Staubli VAL3: teachPoint1.pgx

public program teachPoint1(string x_sKey, num x_nIndex, num x_nPointIndex)
  local num l_nFrameIndex
  local num l_nToolIndex
  local frame l_fFrame
  local tool l_tTool
  local bool l_bResult
  local pointRx l_pPoint
begin
  link(l_tTool,flange)
  link(l_fFrame,world)
  //  l_bResult=userPageConfirm("是否记录当前点位："+toString("",x_nIndex))
  //  if l_bResult
  l_nFrameIndex=trajTemp:tTrajItem[x_sKey].nFrameIndex
  l_nToolIndex=trajTemp:tTrajItem[x_sKey].nToolIndex
  call savedata:getFrame(l_nFrameIndex,l_fFrame)
  call savedata:getTool(l_nToolIndex,l_tTool)


  trajTemp:tTrajItem[x_sKey].pPointItem[x_nIndex].jJointRx=herej()
  l_pPoint=jointToPoint(l_tTool,l_fFrame,herej())
  switch x_nPointIndex
    case 0
      trajTemp:tTrajItem[x_sKey].pPointItem[x_nIndex].pInter.trsf=l_pPoint.trsf
      trajTemp:tTrajItem[x_sKey].pPointItem[x_nIndex].pInter.config=l_pPoint.config
    break
    case 1
      trajTemp:tTrajItem[x_sKey].pPointItem[x_nIndex].pPointRx.trsf=l_pPoint.trsf
      trajTemp:tTrajItem[x_sKey].pPointItem[x_nIndex].pPointRx.config=l_pPoint.config
    break
  endSwitch

  //x_bToSave=true
  //  endIf
end
